{attribute 'qualified_only'}
{attribute 'strict'}
{attribute 'to_string'}
TYPE E_LogRecordExporterFailureReason :
(
	NA := 0,  // No failure occurred.
	ACTIVE_EXPORT_IN_PROGRESS,  // The exporter cannot accept another batch while an export is active.
	QUEUE_TRANSFER_FAILURE,  // Records could not be transferred into the exporter queue.
	SERIALIZATION_FAILURE,  // The accepted records could not be serialized.
	BUFFER_ALLOCATION_FAILURE,  // The serialized payload buffer could not be allocated.
	FILE_OPEN_FAILURE,  // The destination file could not be opened.
	FILE_WRITE_FAILURE,  // The serialized payload could not be written.
	FILE_CLOSE_FAILURE,  // The destination file could not be closed.
	HTTP_URL_PARSE_FAILURE,  // The configured endpoint URL could not be parsed.
	HTTP_REQUEST_FAILURE,  // The HTTP request could not be sent or completed.
	HTTP_STATUS_FAILURE  // The server responded with a non-success HTTP status code.
) UDINT;
END_TYPE

(* stored: Version 1.1.0.1
   EnumerationTextList E_LogRecordExporterFailureReason: Id {e1d90d84-b23a-4a95-a760-813f7018766a} *)
